Staubli VAL3: utAppearance.dtx

public string sBackgroundColour
public string sBackgroundImage
public string sColour
public bool bVisibility
